Yaskawa INFORM job: PRECPRO.JBI

/JOB
//NAME PRECPRO
//POS
///NPOS 6,0,0,0,0,0
///TOOL 9
///POSTYPE PULSE
///PULSE
C00000=22262,-88873,99586,-534,455,101283
C00001=22262,-88873,99586,-534,455,101283
C00002=-22261,88872,-99584,534,0,-101283
C00003=-22261,88872,-99584,534,0,-101283
C00004=-22261,88872,-99584,534,0,-101283
C00005=22262,-88873,99586,-534,455,101283
//INST
<volatile>
///COMM Generated using RoboDK
///ATTR SC,RW
///GROUP1 RB1
NOP
'Program generated by RoboDK v
'6.0.7 for Yaskawa Motoman DX1
'350D on XX/XX/XXXX 18:00:00
'Using nominal kinematics.
'Using Frame P (targets wrt ba
'se):
'0.0,-0.0,1000.0,90.0,-0.5,0.1
'Tool Tool P should be close t
'o:
'0.1,-0.4,123.5,-45.2,0.0,0.0
MOVJ C00000 VJ=50.00
MOVL C00001 V=100.0
MOVL C00002 V=100.0
MOVJ C00003 VJ=50.00
MOVJ C00004 VJ=50.00
TIMER T=0.00
TIMER T=1.00
MOVL C00005 V=66.7
END
